(*
	Processor test double that writes each emitted record's string body to the TwinCAT ADS log
	(the Error List) instead of exporting it. Stage it in place of a real processor to watch records
	arrive during manual debugging; no automated test asserts on its output.
*)
FUNCTION_BLOCK FB_LogRecordProcessor_ConsolePrinter EXTENDS FB_LogRecordProcessor_Simple

METHOD onEmit
VAR_INPUT
	logRecord: REFERENCE TO FB_LogRecord;
END_VAR
THIS^.writeToConsole(logRecord);
END_METHOD

METHOD writeToConsole
VAR_INPUT
	logRecord: REFERENCE TO FB_LogRecord;
END_VAR
VAR
	body: POINTER TO FB_String;
END_VAR
IF logRecord.body <> 0 AND_THEN logRecord.body^.eType = E_ValueType.E_String THEN
	body := logRecord.body;
	ADSLOGSTR(
		ADSLOG_MSGTYPE_ERROR,
		body^.pString^,
		''
	);
END_IF
END_METHOD

END_FUNCTION_BLOCK

(* stored: Version 1.1.0.1
   POU FB_LogRecordProcessor_ConsolePrinter: Id {fbf4b219-b8fc-4773-8575-46cdfadab41e}, SpecialFunc None
   Method onEmit: Id {9f76947b-2126-437d-8b6c-01496aeeff5f}
   Method writeToConsole: Id {72e1877d-8ae1-4395-b68e-02541697117a} *)
